Universal Robots PolyScope program: ex03_program_test.urp

Program ex03_program_test (installation=safety_included directory=/ursim/programs createdIn=5.9.4.1031232 lastSavedIn=5.9.4.1031232 robotSerialNumber=20195599999)
Calibrated DH parameters: a=[0, -0.425, -0.3922, 0, 0, 0]; d=[0.1625, 0, 0, 0.1333, 0.0997, 0.0996]; alpha=[1.570796, 0, 0, 1.570796, -1.570796, 0]; deltaTheta=[0, 0, 0, 0, 0, 0]
Robot Program (runOnlyOnce=false)
  SafeHome (positionOptionType=SPEED_AND_ACCELERATION speed=1.047198 acceleration=1.396263 nextMotionTime=2)
  MoveJ speed 60 deg/s, acceleration 80 deg/s^2 (useActiveTCP=true) feature=Base
    Waypoint Waypoint_1: TCP in base x=-212.52 y=-93.239 z=250.867 mm, rx=-0.8971 ry=-2.5364 rz=-0.5614 rad; joints [-109.071, -50.638, -146.354, -97.676, 68.137, 24.721] deg
  Popup Message (haltProgram=false message=Moved to position Waypoint_1 inputType=Text)
